# EPICS autosave request: iocs/mca-amptek-ioc/db/Amptek_settings.req
$(P)$(R)InputPolarity
$(P)$(R)Clock
$(P)$(R)Gain
$(P)$(R)Gate
$(P)$(R)PeakingTime
$(P)$(R)FastPeakingTime
$(P)$(R)FlatTopTime
$(P)$(R)SlowThreshold
$(P)$(R)FastThreshold
$(P)$(R)PUREnable
$(P)$(R)MCASource
$(P)$(R)ConfigFileName
$(P)$(R)ReadStatus.SCAN
$(P)$(R)SetDetTemp
$(P)$(R)SetHighVoltage
$(P)$(R)MCSLowChannel
$(P)$(R)MCSHighChannel
$(P)$(R)AuxOut1
$(P)$(R)AuxOut2
$(P)$(R)AuxOut34
$(P)$(R)Connector1
$(P)$(R)Connector2
$(P)$(R)SCAOutputWidth
